(* IEC 61131-3 sources: SortJet_MasterSPS_Aufbau.fbsproj/09_Station/Shuttle/[151,152] Transfershuttle, 2 files *)

(* ---- Transfershuttle_FB_V01_00_00.fb.st ---- *)
(* METADATA
{
	"v3Meta": {
		"objectGuid": "6b86eeab-fdc2-4247-b783-cb86ac5f0d72"
	}
}
*)
FUNCTION_BLOCK Transfershuttle_FB_V01_00_00
VAR_IN_OUT

  // STRUKT
  BasisStationsParameter : StationBasisParameter_ST;

END_VAR
VAR_INPUT

  // BOOLEAN
  bpStarteSpeicherfachValidierung       : BOOL;
  bpTransfershuttleVerbundAktiv         : BOOL := false; // Hinweis: Transferverbund zwischen 2 Transvershuttle-Systmen aktiv
  bpScheibenNeuAusrichten               : BOOL;

  // REAL
  rpVorpositionierweg                   : REAL; // Auftragsdaten: Der Weg der Vorpositioniert werden soll

  // STRUCT
  stpInTransportVerbund                 : Interface_TransfershuttleVerbund; // STRUKTUR: Schnittstelle zwischen den Transfershuttlen

END_VAR
VAR_OUTPUT

  // BOOLEAN
  bpShuttleKannSicherVerfahrenWerden     : BOOL; // Shuttle kann sicherverfahren werden - Shuttle ist unten , Abfragen sind unten
  bpAnforderungBetriebsstopp             : BOOL; // Hinweis: Anforderung zum setzen des Betriebsstopps fuer die Auslaufseite des Transfershuttles
  bpSpeicherfachValidierungAbgeschlossen : BOOL; // BETRIEBSART: Validierung des Speicherfachs wurde abgeschlossen
  bpScheibenNeuAusrichtenAbgeschlossen   : BOOL;

  // WORD
  wpAusnahmefehlerTyp    : WORD := WORD#0; // Sensorfehlertyp: 0 = Allgemeiner Fehler / 1 = Einlauf / 2 = Auslauf / 3 = Ein- Aus- Lauf

  // DWORD
  dwlHandfunktionen       : DWORD;  // Handfunktionen: 0..31 Bit
  dwpHandfunktionenReturn : DWORD;  // Aktive Handfunktionen, gleiche Bitbelegung wie dwlHandfunktionen

  // INT
  iPhaseSpeichervalidierung : INT;

  // REAL
  rpVorpositionierterWeg          : REAL; // OUT-STATUS: Status wie weit vorpositioniert wurde
  rpIstPositionNachPositionierung : REAL;

  // ENUM
  ReservierungsStatus    : TransfershuttleReservierungsTyp_EN;

  // STRUKTUR
  stpOutTransportVerbund : Interface_TransfershuttleVerbund; // STRUKTUR: Schnittstelle zwischen den Transfershuttlen

END_VAR
VAR

  // Rueckmeldung der Handfunktionen zum MMI
  dwlHandfunktionenZuletztGesendet           : DWORD;

  // BOOLEAN
  blErsterZyklus                             : BOOL := TRUE; // Initialisierung
  blZielPositionErreicht                     : BOOL;
  blShuttleKannSicherVerfahrenWerden         : BOOL := FALSE;
  blUpdateTimer                              : BOOL; // VERFAHRLOGIK
  blValidierungLuftabfrageAuslaufUnten       : BOOL := FALSE;
  blValidierungLuftabfrageEinlaufUnten       : BOOL := FALSE;
  blHinweisGenerierenSKAusgeloest            : BOOL := FALSE;

  // WORD
  wlWatchIONachrichtenNummer                 : WORD;

  // STEPS
  steplEintransport          : Steps_TE;
  steplAustransport          : Steps_TE;
  steplVortransport          : Steps_TE;
  steplReset                 : Steps_TE;
  steplCheck                 : Steps_TE;
  steplReferenz              : Steps_TE;
  steplVorabpositionierung   : Steps_TE;
  steplScheibenNeuAusrichten : Steps_TE;

  // TRIGGER
  ftlBausteinDeaktivierung   : F_TRIG;

  // TIMER
  tonlMaxWarteAufResetErfolgreich     : TON;
  tonlUpdateTimer                     : TON;
  tonlWarteShuttleSicherVerfahren     : TON; // Max. Warte Zeit wenn Shuttle nicht verfahren koennte, damit die WatchIO vorher aufkommen koennen *)

  // BAUSTEINE
  Glastransport                   : Transfershuttle_Glastransport_FB_V01_00_00;
  Zentralschmierung               : Zentralschmierung_DLS_4xxi_FB_V01_00_00;
  Querfahrt                       : Querfahrt_Shuttle_FB_V01_00_00;

END_VAR

VAR

  // HARDWARE - EINGAENGE
  in_bSensorShuttleOben                                       : BOOL;
  in_bSensorShuttleUnten                                      : BOOL;
  in_bSensorScheibenKontrolleAuslaufSeiteOben                 : BOOL;
  in_bSensorScheibenKontrolleAuslaufSeiteUnten                : BOOL;
  in_bSensorScheibenKontrolleAuslaufSeiteFrei                 : BOOL; // Öffner
  in_bSensorScheibenKontrolleEinlaufSeiteOben                 : BOOL;
  in_bSensorScheibenKontrolleEinlaufSeiteUnten                : BOOL;
  in_bSensorScheibenKontrolleEinlaufSeiteFrei                 : BOOL; // Öffner
  in_bDruckluftEinlaufSeiteOK                                 : BOOL;
  in_bDruckluftAuslaufSeiteOK                                 : BOOL;
  in_bDruckluftWartungseinheitOK                       AT %I* : BOOL;
  in_bLeitungsschutz_Querfahrt_OK                      AT %I* : BOOL;

END_VAR

//-------------------------------------------------------------------------------------------------
// INITIALISIERUNG
//-------------------------------------------------------------------------------------------------
IF ( blErsterZyklus ) THEN
  blErsterZyklus:=FALSE;

  A_Baustein_Initialisierung();

END_IF

in_bSensorScheibenKontrolleEinlaufSeiteFrei := Glastransport.Antrieb.blSensoren[1];
in_bSensorScheibenKontrolleAuslaufSeiteFrei := Glastransport.Antrieb.blSensoren[2];

//-------------------------------------------------------------------------------------------------
// DEAKTIVIERUNG
//-------------------------------------------------------------------------------------------------

(* Hinweis:
   - Werte wieder passend abloeschen, wenn der Baustein wieder aktiviert wird
*)
ftlBausteinDeaktivierung( CLK := BasisStationsParameter.stMKs.bDeaktivieren );

IF ( ftlBausteinDeaktivierung.Q ) THEN

  SendShuttlePosition();

  BasisStationsParameter.bEintransportAbgeschlossen[cWAND_1] := FALSE;
  BasisStationsParameter.bAustransportAbgeschlossen[cWAND_1] := FALSE;
  BasisStationsParameter.bVortransportAbgeschlossen[cWAND_1] := FALSE;
  BasisStationsParameter.bVorabpositionierenAbgeschlossen    := FALSE;
  bpSpeicherfachValidierungAbgeschlossen := FALSE;
  bpScheibenNeuAusrichtenAbgeschlossen   := FALSE;

  BasisStationsParameter.bIstReferenziert       := FALSE;
  BasisStationsParameter.bCheckAbgeschlossen    := FALSE;
  BasisStationsParameter.bReferenzAbgeschlossen := FALSE;

END_IF

(* Hinweis:
   - Deaktivierung des Bausteins
     => Der Baustein wird zum Ende der RETURN-Anweisung verlassen
*)
IF ( BasisStationsParameter.stMKs.bDeaktivieren ) THEN

  IF ( apgTransfershuttleVerfahrparameter[BasisStationsParameter.stMKs.stStationsNummern.NummerSPS].eParkposition = PARKPOSITION_MAX ) THEN
    BasisStationsParameter.rAktuellePositionQuerfahrt := apgTransfershuttleVerfahrparameter[BasisStationsParameter.stMKs.stStationsNummern.NummerSPS].rParkpositionMaximum;
  ELSE
    BasisStationsParameter.rAktuellePositionQuerfahrt := apgTransfershuttleVerfahrparameter[BasisStationsParameter.stMKs.stStationsNummern.NummerSPS].rParkpositionMinimum;
  END_IF

  BasisStationsParameter.bEintransportAbgeschlossen[cWAND_1] := TRUE;
  BasisStationsParameter.bAustransportAbgeschlossen[cWAND_1] := TRUE;
  BasisStationsParameter.bVortransportAbgeschlossen[cWAND_1] := TRUE;
  BasisStationsParameter.bVorabpositionierenAbgeschlossen    := TRUE;
  BasisStationsParameter.bReset                              := FALSE;
  bpSpeicherfachValidierungAbgeschlossen := TRUE;
  bpScheibenNeuAusrichtenAbgeschlossen   := TRUE;

  BasisStationsParameter.bIstReferenziert       := TRUE;
  BasisStationsParameter.bCheckAbgeschlossen    := TRUE;
  BasisStationsParameter.bReferenzAbgeschlossen := TRUE;

  BasisStationsParameter.bFehler                := FALSE;
  BasisStationsParameter.wFehlerNummer          := cMELDUNG_NULL;

  HandfunktionenStatus();
  RETURN;

END_IF

//-------------------------------------------------------------------------------------------------
// AKTIONEN
//-------------------------------------------------------------------------------------------------

(* Hinweis:
   - SystemCheck
*)
Systemcheck();

(* Hinweis:
   - Automatik- Aktionen
*)
Eintransport();
Vortransport();
Austransport();
Vorabpositionierung();
//Transportkopplung();
ScheibenNeuAusrichten();

(* Hinweis:
   - Gesonderte- Aktionen
*)
SpeicherfachValidierung();

(* Hinweis:
   - Basis- Aktionen
*)

Reset();
Referenz();
Handfunktionen();
Meldungen();

A_Schnittstelle();
A_Aufrufe();
A_Ausgaenge();
END_FUNCTION_BLOCK

(* ---- Transfershuttle_Glastransport_FB_V01_00_00.fb.st ---- *)
(* METADATA
{
	"v3Meta": {
		"objectGuid": "2254a377-1dbb-47e5-a6cb-497511b1e2ee"
	}
}
*)
FUNCTION_BLOCK Transfershuttle_Glastransport_FB_V01_00_00
VAR_INPUT

  // BOOLEAN
  bpAktivieren                                       : BOOL;
  bpEintransport                                     : BOOL;
  bpAustransport                                     : BOOL;
  bpVortransport                                     : BOOL;
  bpFahreReferenz                                    : BOOL;
  bpAutomatikAktiv                                   : BOOL;
  bpSlaveKopplung                                    : BOOL;
  bpCheck                                            : BOOL;
  bpReset                                            : BOOL;
  bpShuttleVerfaehrt                                 : BOOL;
  bpHand                                             : BOOL;
  bpFreigabe                                         : BOOL;
  bpShuttleAbsenken                                  : BOOL;
  bpHandfahrenPlus                                : BOOL;
  bpHandfahrenMinus                                : BOOL;
  bpHandGlastransportAnheben                         : BOOL;
  bpHandScheibenKontrolleEinlaufseiteAnheben         : BOOL;
  bpHandScheibenKontrolleAuslaufseiteAnheben         : BOOL;
  bpHandScheibenKontrolleEinlaufseiteEin             : BOOL;
  bpHandScheibenKontrolleAuslaufseiteEin             : BOOL;
  bpStarteHebeVorgang                                : BOOL;
  bpRueckwaertsEintransportieren                     : BOOL;
  bpRueckwaertsAustransportieren                     : BOOL;
  bpGlastransportTest                                : BOOL;
  bpSpeicherfachValidierung                          : BOOL; // Betriebsmodus: Speicherfach wird ueberprueft ob beide Luftabfragen frei und somit kein Glas uebersteht
  bpScheibentrennung                                 : BOOL := FALSE;
  bpAnforderungTransportkopplung                     : BOOL := FALSE;
  blSensorGlastransportOben                          : BOOL;
  blSensorGlastransportUnten                         : BOOL;
  bpSensorScheibenKontrolleAuslaufSeiteOben          : BOOL;
  bpSensorScheibenKontrolleAuslaufSeiteUnten         : BOOL;
  bpSensorScheibenKontrolleAuslaufSeiteFrei          : BOOL; // Oeffner
  bpSensorScheibenKontrolleEinlaufSeiteOben          : BOOL;
  bpSensorScheibenKontrolleEinlaufSeiteUnten         : BOOL;
  bpSensorScheibenKontrolleEinlaufSeiteFrei          : BOOL; // Oeffner
  blDruckluftEinlaufSeiteOK                          : BOOL;
  blDruckluftAuslaufSeiteOK                          : BOOL;
  bpTransfershuttleVerbundAktiv                      : BOOL := FALSE; // Hinweis: Transferverbund zwischen 2 Transvershuttle aktiv
  bpOptionSensorEinlauf                              : BOOL := TRUE;  // Hinweis: Option ob der Sensorvorhanden ist
  bpOptionSensorAuslauf                              : BOOL := TRUE;  // Hinweis: Option ob der Sensorvorhanden ist
  bpScheibenNeuAusrichten                            : BOOL;
  bpOptionTransfershuttleMitFaecherwagen             : BOOL;
  bpOptionTransfershuttleMitUltraschallSensoren      : BOOL;
  bpOptionMasterSlaveAustransport                    : BOOL;
  bpOptionTransfershuttleFaecherwagenKurzeScheibenTieferEintransportieren : BOOL; // Debug-Funktion: wird nur von Hand (Online) gesetzt, kurze Scheiben 150 mm tiefer eintransportieren

  // REAL
  rpVorpositionierweg : REAL; // Auftragsdaten: Der Weg der Vorpositioniert werden soll

  // STRUCT
  InGlasTransportVorgaenger   : Interface_GlasTransport; // STRUKTUR: Informationen ueber den Aus- Ein- Transport der Vorgaengerstation
  InGlasTransportNachfolger   : Interface_GlasTransport; // STRUKTUR: Informationen ueber den Aus- Ein- Transport der Nachfolge- Station
  stpInTransportVerbund       : Interface_TransfershuttleVerbund;
  pAuftrag                    : Auftragsdaten_ST;        // AUFTRAG: Aktuelle daten zum Auftrag [Laenge, Hoehe, Modelle]
  pSystemCheckDaten           : Auftragsdaten_ST;        // Hinweis: Daten fuer den SystemCheck
  stMasterSlaveConfig         : MasterSlaveConfig_ST;
  stStationsNummern           : Station_ST;

  // POINTER
  ppParameterBaustein     : REFERENCE TO Parameter_TransfershuttleGlastransport;
  ppAntriebsInformationen : REFERENCE TO AntriebsInformationen;

END_VAR
VAR_OUTPUT

  // BOOLEAN
  bpDone                                 : BOOL;
  bpFehler                               : BOOL;
  bpAktiv                                : BOOL;
  bpSlaveAktiv                           : BOOL;
  bpBereitZumVerfahren                   : BOOL := FALSE;
  bpScheibeFaehrtUeberAuslauf            : BOOL; // Variable zum nehmen der Verfahrfreigabe des Shuttles da Glas in den Verfahrbereich liegen koennte
  bpScheibeFaehrtUeberEinlauf            : BOOL; // Variable zum nehmen der Verfahrfreigabe des Shuttles da Glas in den Verfahrbereich liegen koennte
  bpAnforderungBetriebsstopp             : BOOL; // Hinweis: Anforderung zum setzen des Betriebsstopps fuer die Auslaufseite des Transfershuttles
  bprtScheibe                            : BOOL; // Scheibenzaehler, funktion wie ein Trigger
  bpOutBereitZumAustransport             : BOOL;
  bpOutBereitZumEintransport             : BOOL;
  bpSpeicherfachValidierungAbgeschlossen : BOOL;
  bpSensorEinlauf                        : BOOL; // Sensorik Ausgang: Setzen der Sensorik fuer die Transportkopplung
  bpSensorAuslauf                        : BOOL; // Sensorik Ausgang: Setzen der Sensorik fuer die Transportkopplung

  // WORD
  wpFehlerNr              : Fehlerkonstanten_EN;
  wpAusnahmefehlerTyp     : WORD := WORD#0; // Sensorfehlertyp: 0 = Allgemeiner Fehler / 1 = Einlauf / 2 = Auslauf / 3 = Ein- Aus- Lauf

  // REAL
  rpOutGeschwindigkeit   : REAL; // OUT STATUS: Aktuelle Geschwindigkeit
  rpVorpositionierterWeg : REAL; // OUT STATUS: Beschreibt den Weg der Vorpositioniert wurde

  // STRUCT
  stpOutTransportVerbund : Interface_TransfershuttleVerbund;

END_VAR
VAR

  // BOOLEAN
  blErsterZyklus                               : BOOL := TRUE;
  blBereitZumGlastransport                     : BOOL := FALSE;
  blEinlaufSensor                              : BOOL; // entprellter Eingangssensor
  blAuslaufSensor                              : BOOL; // entprellter Ausgangssensor
  blScheibenMerker                             : BOOL := FALSE; // Scheibe lag nach dem Positionieren noch auf dem Einlaufsensor => Quittung beim Freifahren
  blFehlerAusloesen                            : BOOL; // Hinweis: Es muss ggf ein Fehler ausgeloest werden wenn ein Sensor angefahren und programmgesteuert wieder Freigefahren wurde
  blMeldungAuslaufAbfrageBelegt                : BOOL := FALSE; // Hinweis: Sensorik beim Pruefen belegt
  blMeldungEinlaufAbfrageBelegt                : BOOL := FALSE; // Hinweis: Sensorik beim Pruefen belegt
  blSensorPruefungEinlaufsensorBelegt          : BOOL := FALSE;
  blSensorPruefungAuslaufsensorBelegt          : BOOL := FALSE;
  blAbgeschlossenAustransport                  : BOOL := FALSE;
  blAbgeschlossenEintransport                  : BOOL := FALSE;
  blEintransportDefaultLuftabfrage             : BOOL := FALSE;
  blAustransportDefaultLuftabfrage             : BOOL := FALSE;
  blSchnittstelle_bBereitZumTransportVerbund   : BOOL := FALSE;
  blSchnittstelle_bAnforderungTransportVerbund : BOOL := FALSE;
  blScheibenKontrolleEinlaufseiteEin           : BOOL;
  blScheibenKontrolleAuslaufseiteEin           : BOOL;
  blReduzierteGeschwindigkeit                  : BOOL;

  // WORD
  wlSubIndex : WORD;

  // INT
  ilScheibenZaehler                          : INT; // Scheibenzaehlen

  // REAL
  rlAntriebsPositionBeiStart                 : REAL;
  rlMaxStreckeErsteScheibe                   : REAL; // Max. Weg bis zur ersten Scheibe: Laenge der abgebenden Station, ohne bekannte Laenge die eigene Stationslaenge
  rlAntriebsPositionStartVortransport        : REAL; // Ist-Position beim Start Vortransport fuer rpVorpositionierterWeg
  rlAntriebspositionBeiAuslaufSensorBelegung : REAL;
  rlWegDifferenzNachStopSensorBelegung       : REAL;
  rlPositionScheibenAnfangErkannt            : REAL;
  rlZielPosition                             : REAL;
  rlStreckeBisZurVerzoegerung                : REAL;
  rlGlasgewicht                              : REAL;

  // STEPS
  steplEintransport                   : Steps_TE;
  steplAustransport                   : Steps_TE;
  steplVortransport                   : Steps_TE;
  steplReset                          : Steps_TE;
  steplReferenz                       : Steps_TE;
  steplCheck                          : Steps_TE;
  steplHebeVorgang                    : Steps_TE;
  steplGlastransporttest              : Steps_TE;
  steplSpeicherfachValidierung        : Steps_TE;
  steplEintransportDefaultLuftabfrage : Steps_TE;
  steplAustransportDefaultLuftabfrage : Steps_TE;
  steplSlave                          : Steps_TE;
  steplScheibenNeuAusrichten          : Steps_TE;

  // FLANKEN
  rtriglFehlerAktiv                   : R_TRIG; // Fehler-Bit Triggern
  ftriglAuslaufsensorBelegt           : F_TRIG; // fallende Flanke: Auslaufsensor wurde angefahren
  ftriglEinlaufsensorBelegt           : F_TRIG; // fallende Flanke: Einlaufsensor wurde angefahren

  // TIMER
  tonlGlastransportOben                             : TON;
  tonlAntriebNichtFreigegeben                       : TON;
  tonlUeberwachungSensorFreifahren                  : TON;
  tonlKontrolleEinlaufOben                          : TON;
  tonlKontrolleEinlaufUnten                         : TON;
  tonlKontrolleAuslaufOben                          : TON;
  tonlKontrolleAuslaufUnten                         : TON;
  tonlWartenAufAnheben                              : TON;
  tonlWartenAufSenken                               : TON;
  tonlEinlaufWirklichFrei                           : TON;
  tonlAuslaufWirklichFrei                           : TON;
  tonlEinlaufsensorTesten                           : TON;
  tonlAuslaufsensorTesten                           : TON;
  tonlMaxWarteAufResetErfolgreich                   : TON;
  tonlUberwachungSlaveAktiv                         : TON;
  tonlEinlaufsensorFrei                             : TON; // Luftsensor Einlauf frei, entprellt
  tonlEinlaufsensorBelegt                           : TON; // Luftsensor Einlauf belegt, entprellt
  tonlAuslaufsensorFrei                             : TON; // Luftsensor Auslauf frei, entprellt
  tonlAuslaufsensorBelegt                           : TON; // Luftsensor Auslauf belegt, entprellt
  toflAutoAbschaltung                               : TOF;
  toflAntriebLaeuft                                 : TOF;

  // Antrieb
  Antrieb : REFERENCE TO Rexroth_ctrlX_Drive_Eckelmann_MC_V01_02_02;

END_VAR
VAR

  // HARDWARE - AUSGAENGE
  out_bShuttleAnheben                                        : BOOL;
  out_bScheibenKontrolleEinlaufSeiteAuf                      : BOOL; // AUSGAENGE: Luftabfragen heben/senken
  out_bScheibenKontrolleEinlaufSeiteEinschalten              : BOOL;
  out_bScheibenKontrolleAuslaufSeiteAuf                      : BOOL; // AUSGAENGE: Luftabfragen heben/senken
  out_bScheibenKontrolleAuslaufSeiteEinschalten              : BOOL;

END_VAR
VAR CONSTANT

  // TIME
  cZEIT_SENSORIK_FREIFAHREN           : TIME := T#10s;
  cZEIT_UEBERWACHUNG_ANTRIEBSFREIGABE : TIME := T#5S;
  cZEIT_UEBERWACHUNG_SLAVE_AKTIV      : TIME := T#10s;

END_VAR

//-------------------------------------------------------------------------------------------------
// INITIALISIERUNG
//-------------------------------------------------------------------------------------------------
IF ( blErsterZyklus ) THEN

  IF ( __ISVALIDREF(ppAntriebsInformationen) ) THEN

    blErsterZyklus := FALSE;

    Antrieb REF= pgAntriebe[ppAntriebsInformationen.wAchsID];

    (* Hinweis:
       - Initialisierung Antriebsinformationen
    *)
    Antrieb.ppAntriebsInformationen REF= ppAntriebsInformationen;

    (* Hinweis:
       - Für die Zielpunktkontrolle muss im ersten Zyklus die Zielposition initialisiert werden
    *)
    Antrieb.rpZielPosition := Antrieb.rpIstPosition;

    (* Hinweis:
       - Antriebswerte vorinitialisieren
    *)
    Antrieb.rpGeschwindigkeit := ppAntriebsInformationen.rpMaxGeschwindigkeit;
    Antrieb.rpBeschleunigung  := ppAntriebsInformationen.rpMaxBeschleunigung;
    Antrieb.rpVerzoegerung    := ppAntriebsInformationen.rpMaxVerzoegerung;
    Antrieb.rpRuckzeit        := ppAntriebsInformationen.rpMaxRuckzeit;

  ELSE
    RETURN;
  END_IF

END_IF

//-------------------------------------------------------------------------------------------------
// DEAKTIVIEREN
//-------------------------------------------------------------------------------------------------
IF ( NOT bpAktivieren ) THEN

  bpDone := TRUE;

  (* Hinweis:
     - Ausnahmesituationen
  *)
  bpFehler   := FALSE;
  wpFehlerNr := cMELDUNG_NULL;

  RETURN;

END_IF

//-------------------------------------------------------------------------------------------------
// BAUSTEIN: SCHNITTSTELLE
//-------------------------------------------------------------------------------------------------
(* Hinweis:
   - Schnittstelle zwischen den Unterflur-Shuttle wenn diese zusammen arbeiten sollen
*)
stpOutTransportVerbund.wpMmiNummer                  := stStationsNummern.NummerSPS;
stpOutTransportVerbund.bEinlaufsensor               REF= bgFALSE;
stpOutTransportVerbund.bAuslaufsensor               REF= bgFALSE;
stpOutTransportVerbund.bMasterSlaveVerbundAktiv     REF= bpSlaveAktiv; // Slave ist mit dem Master gekoppelt
stpOutTransportVerbund.bBereitZumTransportVerbund   REF= blSchnittstelle_bBereitZumTransportVerbund;
stpOutTransportVerbund.bAnforderungTransportVerbund REF= blSchnittstelle_bAnforderungTransportVerbund;
stpOutTransportVerbund.rGeschwindigkeit             REF= rpOutGeschwindigkeit;
stpOutTransportVerbund.bFehler                      REF= bpFehler;

//-------------------------------------------------------------------------------------------------
// BAUSTEIN: SENSOREN \ TIMER \ GESCHWINDIGKEITEN \ ETC.
//-------------------------------------------------------------------------------------------------
// [TIMER] Allgemein:
toflAntriebLaeuft(IN:=Antrieb.bpAntrieblaeuft, PT := T#350MS);

// [TIMER] Kontrolle Sensoren:
//   - Glastransport Oben
tonlGlastransportOben(IN := blSensorGlastransportOben, PT := t#500ms);

// ---------------------------------------------------------------------------------------
//  TRANSFERSHUTTLE MIT EINEM LUFTABFRAGEN TYP
//
//  Hinweis:
// - n/c
// ---------------------------------------------------------------------------------------

// LUFTABFRAGEN [3- 12 MM]
//   - [TIMER] Kontrolle Sensoren:
//     => Einlauf- Sensoren [ Luftsenoren] Frei | Belegt
//     => Auslauf- Sensoren [ Luftsenoren] Frei | Belegt
//     => frei und belegt werden beide entprellt (50 ms), Scheibenzaehlung erst bei sicher freiem Sensor
tonlEinlaufsensorFrei(IN:= bpSensorScheibenKontrolleEinlaufseiteFrei, PT := t#50ms);
tonlEinlaufsensorBelegt(IN:= NOT bpSensorScheibenKontrolleEinlaufseiteFrei, PT := t#50ms);
tonlAuslaufsensorFrei(IN:= bpSensorScheibenKontrolleAuslaufSeiteFrei, PT := t#50ms);
tonlAuslaufsensorBelegt(IN:= NOT bpSensorScheibenKontrolleAuslaufSeiteFrei, PT := t#50ms);

// LUFTABFRAGEN [3- 12 MM]
//   - [TIMER] Kontrolle Sensoren:
//     => Einlauf- Sensoren [ Luftsenoren] Unten | Oben
//     => Auslauf- Sensoren [ Luftsenoren] Unten | Oben
tonlKontrolleEinlaufUnten(IN := bpSensorScheibenKontrolleEinlaufseiteUnten, PT := T#500MS);
tonlKontrolleEinlaufOben(IN := bpSensorScheibenKontrolleEinlaufseiteOben, PT := T#500MS);

tonlKontrolleAuslaufUnten(IN := bpSensorScheibenKontrolleAuslaufseiteUnten, PT := T#500MS);
tonlKontrolleAuslaufOben(IN := bpSensorScheibenKontrolleAuslaufseiteOben, PT := T#500MS);

// LUFTABFRAGEN [3- 12 MM]
//   - Sensorik freifahren
tonlEinlaufWirklichFrei(IN:= NOT blEinlaufsensor, PT := t#500ms);
tonlAuslaufWirklichFrei(IN:= NOT blAuslaufsensor, PT := t#500ms);

// LUFTABFRAGEN [3- 12 MM]
//   - Sensoren:
//     => Einlauf / Auslauf
blEinlaufsensor := tonlEinlaufsensorBelegt.Q AND ( blDruckluftEinlaufSeiteOK OR bpOptionTransfershuttleMitUltraschallSensoren );
blAuslaufsensor := tonlAuslaufsensorBelegt.Q AND ( blDruckluftAuslaufSeiteOK OR bpOptionTransfershuttleMitUltraschallSensoren );

(* Hinweis [3- 12 MM]:
   - Abfrage ob die Station bereit fuer den Glastransport ist
*)
blBereitZumGlastransport := (    tonlGlastransportOben.Q
                              AND tonlKontrolleEinlaufOben.Q
                              AND ( blDruckluftAuslaufSeiteOK OR bpOptionTransfershuttleMitUltraschallSensoren )
                              AND tonlKontrolleAuslaufOben.Q
                              AND ( blDruckluftEinlaufSeiteOK OR bpOptionTransfershuttleMitUltraschallSensoren ) );

//-------------------------------------------------------------------------------------------------
// BAUSTEIN: AKTIONEN
//-------------------------------------------------------------------------------------------------
(* Hinweis:
   - Aktion zur Abhandlung von Transfershuttle mit nur einer physikalisch verbauten
     Luftabfrage
*)
Steuerung_OptionaleLuftabfragen();

(* Hinweis:
   - Aufruf der Aktion SystemCheck
   - Starten des SystemChecks mittels Riemen
*)
Systemcheck();

// Aktion [Automatik]:
//   - Starten der Automatik- Aktionen
//     => Eintransport
//     => Austransport
//     => etc.
Eintransport();
Eintransport_Default_Luftabfrage();

Austransport();
Austansport_Default_Luftabfrage();

SlaveBetrieb();

HebeVorgang();

SpeicherTest();

SpeicherfachValidierung();

Vortransport();

ScheibenNeuAusrichten();

// Aktion[Basis]:
//   - Basis Bausteinaktionen
Reset();
Referenz();
Meldungen();
Handfunktionen();
SteuerungLuftschranken();

//-------------------------------------------------------------------------------------------------
// BAUSTEIN: VORTRANSPORT [SPEICHER]
//-------------------------------------------------------------------------------------------------
IF ( bpShuttleAbsenken ) THEN
  out_bShuttleAnheben := FALSE;
  out_bScheibenKontrolleAuslaufSeiteAuf := FALSE;
  blScheibenKontrolleAuslaufseiteEin    := FALSE;
  out_bScheibenKontrolleEinlaufSeiteAuf := FALSE;
  blScheibenKontrolleEinlaufseiteEin    := FALSE;

  bpShuttleAbsenken := FALSE;
END_IF

//-------------------------------------------------------------------------------------------------
// BAUSTEIN: ZUWEISUNGEN UND AUFRUFE
//-------------------------------------------------------------------------------------------------
// Glastransportfreigabe
toflAutoAbschaltung( IN := (  bpAutomatikAktiv
                             AND ( bpEintransport
                                   OR bpAustransport
                                   OR bpStarteHebeVorgang
                                   OR bpVortransport))
                     OR bpCheck
                     OR bpSlaveKopplung
                     OR bpSpeicherfachValidierung
                     OR bpScheibenNeuAusrichten
                     OR bpHandfahrenPlus
                     OR bpHandfahrenMinus
                     OR bpFahreReferenz,
                     PT:=( WORD_TO_TIME(ppParameterBaustein.wEnergieSparZeit)*1000) );

Antrieb.bpFreigabe            := toflAutoAbschaltung.Q AND bpFreigabe;
Antrieb.stStationsNummern     := stStationsNummern;
Antrieb.rpRuckzeit            := ppAntriebsInformationen.rpMaxRuckzeit;

//-------------------------------------------------------------------------------------------------
// BAUSTEIN: AUSGAENGE
//-------------------------------------------------------------------------------------------------

// VERFAHRFREIGABE [3- 12 MM]:
// - Bit ob das Transfershuttle verfahren darf
bpBereitZumVerfahren := (     blSensorGlastransportUnten
                          AND NOT blSensorGlastransportOben
                          AND tonlKontrolleEinlaufUnten.Q
                          AND NOT bpSensorScheibenKontrolleEinlaufseiteOben
                          AND tonlKontrolleAuslaufUnten.Q
                          AND NOT bpSensorScheibenKontrolleAuslaufseiteOben );

// Ausgaeng:
//   - Aktuelle Geschwindigkeit des Antriebs
//     -> Soll- Wertkopplung ( Soll-Geschwindigkeit des Antriebs)
//     -> Ist- Wertkopplung ( Soll-Geschwindigkeit des Antriebs)
IF  ( ( bpEintransport OR bpRueckwaertsEintransportieren ) AND bpOutBereitZumEintransport )
    OR ( bpCheck AND bpOutBereitZumEintransport )
THEN
  rpOutGeschwindigkeit := Antrieb.rpGeschwindigkeit;
ELSE
  rpOutGeschwindigkeit := Antrieb.rpIstGeschwindigkeit;
END_IF

// Ausgaenge:
//   - Sensorik als out-Variablen bereitstellen
//     => Uebergabe der Werte fuer die Transportkopplung (Stationsinterface)
bpSensorEinlauf := blEinlaufSensor;
bpSensorAuslauf := blAuslaufSensor;

// Glastransport [Transfershuttle] arbeitet oder ist gehoben
//   - in Progress
bpAktiv := (   bpEintransport
             OR bpAustransport
             OR bpVortransport
             OR bpSlaveKopplung
             OR bpScheibenNeuAusrichten
             OR bpStarteHebeVorgang
             OR bpCheck
             OR bpDone );

//-------------------------------------------------------------------------------------------------
// BAUSTEIN: FEHLERNUMMER GENERIEREN BEI EINEM TRANSFERSHUTTLE- FEHLER
//-------------------------------------------------------------------------------------------------
(* Hinweis:
   - Ausnahmesituation
*)
rtriglFehlerAktiv(CLK := bpFehler );

IF ( rtriglFehlerAktiv.Q ) THEN

  CASE wpFehlerNr OF

      cMELDUNG_SENSOR_EINLAUF_BELEGT,
        cMELDUNG_AUSTRANSPORT_SENSOR_EINLAUF_BELEGT,
        cMELDUNG_EINTRANSPORT_SENSOR_EINLAUF_BELEGT,
        cMELDUNG_EINTRANSPORT_SENSOR_EINLAUF_NICHT_FREI,
        cMELDUNG_AUSTRANSPORT_SENSOR_EINLAUF_NICHT_FREI:
      wpAusnahmefehlerTyp  := cAUSNAHMESITUATION_EINLAUFSENSOR;

      cMELDUNG_SENSOR_AUSLAUF_BELEGT,
        cMELDUNG_EINTRANSPORT_SENSOR_AUSLAUF_BELEGT,
        cMELDUNG_EINTRANSPORT_SENSOR_AUSLAUF_NICHT_FREI,
        cMELDUNG_AUSTRANSPORT_SENSOR_AUSLAUF_BELEGT,
        cMELDUNG_AUSTRANSPORT_SENSOR_AUSLAUF_NICHT_FREI,
        cMELDUNG_EINTRANSPORT_SENSOR_EINLAUF_ODER_AUSLAUF_BELEGT_FREIFAHREN:
      wpAusnahmefehlerTyp := cAUSNAHMESITUATION_AUSLAUFSENSOR;

      cMELDUNG_SENSOR_EINLAUF_UND_AUSLAUF_BELEGT,
        cMELDUNG_EINTRANSPORT_SENSOR_EINLAUF_UND_AUSLAUF_BELEGT,
        cMELDUNG_AUSTRANSPORT_SENSOR_EINLAUF_UND_AUSLAUF_BELEGT:
      wpAusnahmefehlerTyp := cAUSNAHMESITUATION_EINLAUF_AUSLAUF_SENSOR;

    ELSE
      wpAusnahmefehlerTyp := cAUSNAHMESITUATION_KEIN_SENSOR;

  END_CASE

END_IF

//-------------------------------------------------------------------------------------------------
// BAUSTEIN: SICHERHEIT
//-------------------------------------------------------------------------------------------------
(* Anmerkung:
   - Sollte eine Fahrt anstehen duerfen Glastransport und Luftabfragen nicht angehoben werden!
     [Doppelte Sicherheit ]
*)
out_bScheibenKontrolleAuslaufSeiteAuf := out_bScheibenKontrolleAuslaufSeiteAuf AND NOT bpShuttleVerfaehrt;
out_bScheibenKontrolleEinlaufSeiteAuf := out_bScheibenKontrolleEinlaufSeiteAuf AND NOT bpShuttleVerfaehrt;

out_bShuttleAnheben := out_bShuttleAnheben AND NOT bpShuttleVerfaehrt;
END_FUNCTION_BLOCK
